Omron Sysmac Studio project AutomatedSortingSystem (Sysmac Studio 1.64.0.64008, StandardProject)

# Controller new_Controller_0: NJ301-1100 version 1.69
Units and slaves: Power Supply : NJ-Px3001; CPU : NJ301-1100
Task PrimaryTask (priority 4, period or condition 1000): PRG_SortingSystem

TYPE ST_MotorSimulation : STRUCT
    Enable : BOOL;
    Start : BOOL;
    Stop : BOOL;
    Fault : BOOL;
    RunFeedback : BOOL;
    ResetFault : BOOL;
    MotorRun : BOOL;
    MotorFault : BOOL;
    StartupFault : BOOL;
    FeedbackLostFault : BOOL;
END_STRUCT END_TYPE
TYPE ST_CylinderSimulation : STRUCT
    Enable : BOOL;
    ExtendCmd : BOOL;
    RetractCmd : BOOL;
    SensorExtended : BOOL;
    SensorRetracted : BOOL;
    ResetFault : BOOL;
    ValveExtend : BOOL;
    ValveRetract : BOOL;
    CylinderFault : BOOL;
    ExtendTimeoutFault : BOOL;
    RetractTimeoutFault : BOOL;
END_STRUCT END_TYPE
TYPE ST_SortingSimulation : STRUCT
    AutoMode : BOOL;
    Start : BOOL;
    Stop : BOOL;
    Reset : BOOL;
    ProductDetected : BOOL;
    AtSortingPosition : BOOL;
    ProductType : UINT;  (* 1=A, 2=B, 3=C *)
    CycleActive : BOOL;
    CycleComplete : BOOL;
    SystemFault : BOOL;
    ProductAtExit : BOOL;
END_STRUCT END_TYPE

PROGRAM Program0
VAR
    Motor1 : FB_ConveyorMotor;
    MotorSim : ST_MotorSimulation;
    CylinderSim : ST_CylinderSimulation;
    Cylinder1 : FB_PneumaticCylinder;
END_VAR

(* Section Section0: ladder, written here as Structured Text *)

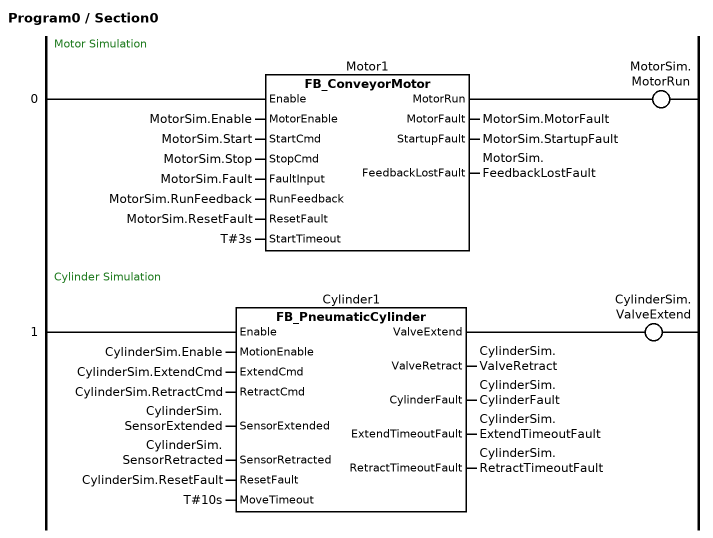
(* Rung 0: Motor Simulation *)
Motor1(Enable := TRUE, MotorEnable := MotorSim.Enable, StartCmd := MotorSim.Start, StopCmd := MotorSim.Stop, FaultInput := MotorSim.Fault, RunFeedback := MotorSim.RunFeedback, ResetFault := MotorSim.ResetFault, StartTimeout := T#3s, MotorFault => MotorSim.MotorFault, StartupFault => MotorSim.StartupFault, FeedbackLostFault => MotorSim.FeedbackLostFault);
MotorSim.MotorRun := Motor1.MotorRun;
(* Rung 1: Cylinder Simulation *)
Cylinder1(Enable := TRUE, MotionEnable := CylinderSim.Enable, ExtendCmd := CylinderSim.ExtendCmd, RetractCmd := CylinderSim.RetractCmd, SensorExtended := CylinderSim.SensorExtended, SensorRetracted := CylinderSim.SensorRetracted, ResetFault := CylinderSim.ResetFault, MoveTimeout := T#10s, ValveRetract => CylinderSim.ValveRetract, CylinderFault => CylinderSim.CylinderFault, ExtendTimeoutFault => CylinderSim.ExtendTimeoutFault, RetractTimeoutFault => CylinderSim.RetractTimeoutFault);
CylinderSim.ValveExtend := Cylinder1.ValveExtend;
END_PROGRAM

PROGRAM PRG_SortingSystem
VAR
    Motor_Conv1 : FB_ConveyorMotor;
    Motor_Conv2 : FB_ConveyorMotor;
    Motor_Conv3 : FB_ConveyorMotor;
    Cylinder_A : FB_PneumaticCylinder;
    Cylinder_B : FB_PneumaticCylinder;
    Conv1 : ST_MotorSimulation;
    Conv2 : ST_MotorSimulation;
    Conv3 : ST_MotorSimulation;
    CylA : ST_CylinderSimulation;
    CylB : ST_CylinderSimulation;
    SortingSim : ST_SortingSimulation;
    TestInput : BOOL;
    TestOutput : BOOL;
    SortingSequence : FB_SortingSequence;
    DevicesReady : BOOL;
    AnyDeviceFault : BOOL;
    SortingState : UINT;
    SystemEnable : BOOL;
    CylinderSim_A : FB_CylinderSimulator;
    CylinderSim_B : FB_CylinderSimulator;
    SimulateCylinderAJam : BOOL := False;
    SimulateCylinderBJam : BOOL := False;
    ResetCylinderAPosition : BOOL := False;
    ResetCylinderBPosition : BOOL := False;
    AlarmManager : FB_AlarmManager;
    ActiveAlarmCode : UINT;
    AlarmActiveStatus : BOOL;
END_VAR

(* Section Section0: ladder, written here as Structured Text *)

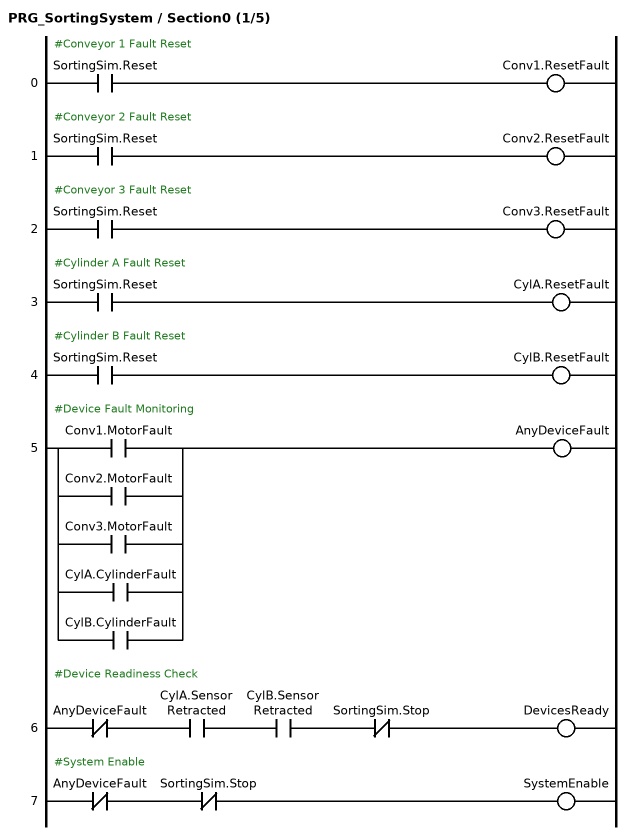
(* Rung 0: #Conveyor 1 Fault Reset *)
Conv1.ResetFault := SortingSim.Reset;
(* Rung 1: #Conveyor 2 Fault Reset *)
Conv2.ResetFault := SortingSim.Reset;
(* Rung 2: #Conveyor 3 Fault Reset *)
Conv3.ResetFault := SortingSim.Reset;
(* Rung 3: #Cylinder A Fault Reset *)
CylA.ResetFault := SortingSim.Reset;
(* Rung 4: #Cylinder B Fault Reset *)
CylB.ResetFault := SortingSim.Reset;
(* Rung 5: #Device Fault Monitoring *)
AnyDeviceFault := Conv1.MotorFault OR Conv2.MotorFault OR Conv3.MotorFault OR CylA.CylinderFault OR CylB.CylinderFault;
(* Rung 6: #Device Readiness Check *)
DevicesReady := NOT AnyDeviceFault AND CylA.SensorRetracted AND CylB.SensorRetracted AND NOT SortingSim.Stop;
(* Rung 7: #System Enable *)
SystemEnable := NOT AnyDeviceFault AND NOT SortingSim.Stop;

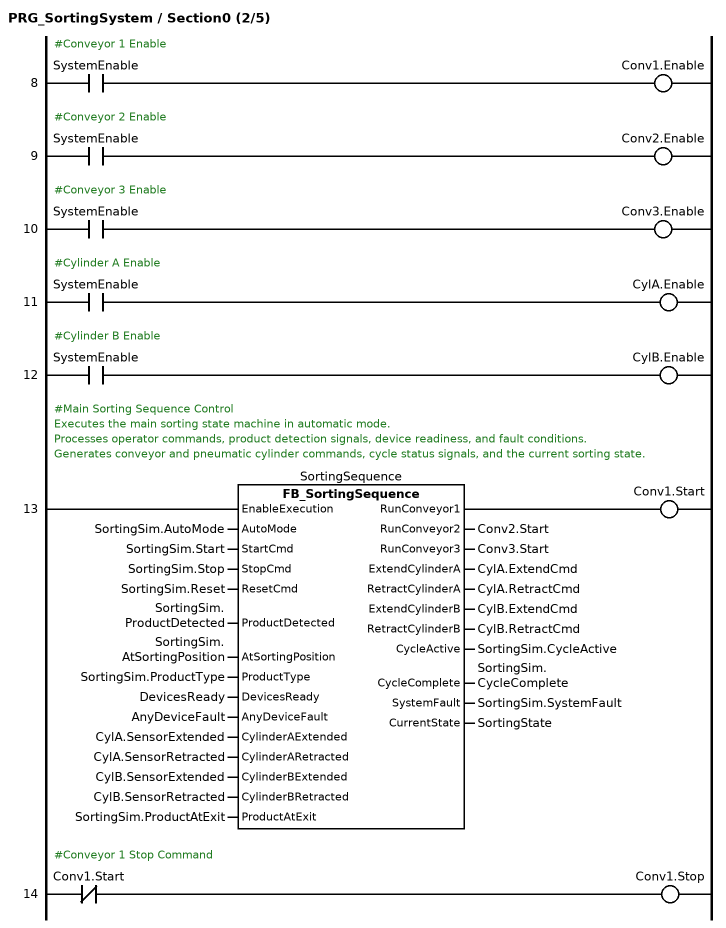
(* Rung 8: #Conveyor 1 Enable *)
Conv1.Enable := SystemEnable;
(* Rung 9: #Conveyor 2 Enable *)
Conv2.Enable := SystemEnable;
(* Rung 10: #Conveyor 3 Enable *)
Conv3.Enable := SystemEnable;
(* Rung 11: #Cylinder A Enable *)
CylA.Enable := SystemEnable;
(* Rung 12: #Cylinder B Enable *)
CylB.Enable := SystemEnable;
(* Rung 13: #Main Sorting Sequence Control / Executes the main sorting state machine in automatic mode. / Processes operator commands, product detection signals, device readiness, and fault conditions. / Generates conveyor and pneumatic cylinder commands, cycle status signals, and the current sorting state. *)
SortingSequence(EnableExecution := TRUE, AutoMode := SortingSim.AutoMode, StartCmd := SortingSim.Start, StopCmd := SortingSim.Stop, ResetCmd := SortingSim.Reset, ProductDetected := SortingSim.ProductDetected, AtSortingPosition := SortingSim.AtSortingPosition, ProductType := SortingSim.ProductType, DevicesReady := DevicesReady, AnyDeviceFault := AnyDeviceFault, CylinderAExtended := CylA.SensorExtended, CylinderARetracted := CylA.SensorRetracted, CylinderBExtended := CylB.SensorExtended, CylinderBRetracted := CylB.SensorRetracted, ProductAtExit := SortingSim.ProductAtExit, RunConveyor2 => Conv2.Start, RunConveyor3 => Conv3.Start, ExtendCylinderA => CylA.ExtendCmd, RetractCylinderA => CylA.RetractCmd, ExtendCylinderB => CylB.ExtendCmd, RetractCylinderB => CylB.RetractCmd, CycleActive => SortingSim.CycleActive, CycleComplete => SortingSim.CycleComplete, SystemFault => SortingSim.SystemFault, CurrentState => SortingState);
Conv1.Start := SortingSequence.RunConveyor1;
(* Rung 14: #Conveyor 1 Stop Command *)
Conv1.Stop := NOT Conv1.Start;

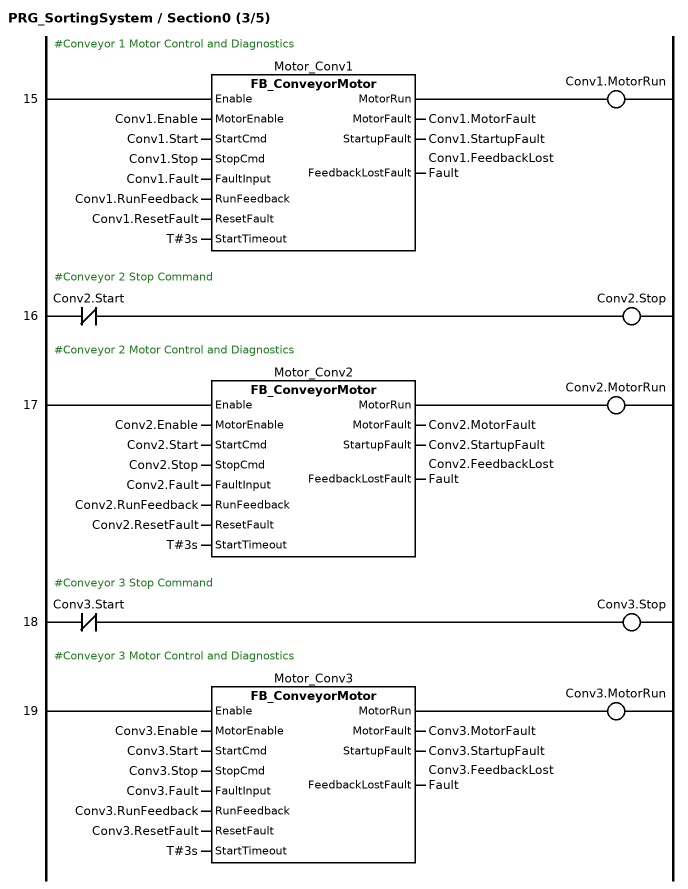
(* Rung 15: #Conveyor 1 Motor Control and Diagnostics *)
Motor_Conv1(Enable := TRUE, MotorEnable := Conv1.Enable, StartCmd := Conv1.Start, StopCmd := Conv1.Stop, FaultInput := Conv1.Fault, RunFeedback := Conv1.RunFeedback, ResetFault := Conv1.ResetFault, StartTimeout := T#3s, MotorFault => Conv1.MotorFault, StartupFault => Conv1.StartupFault, FeedbackLostFault => Conv1.FeedbackLostFault);
Conv1.MotorRun := Motor_Conv1.MotorRun;
(* Rung 16: #Conveyor 2 Stop Command *)
Conv2.Stop := NOT Conv2.Start;
(* Rung 17: #Conveyor 2 Motor Control and Diagnostics *)
Motor_Conv2(Enable := TRUE, MotorEnable := Conv2.Enable, StartCmd := Conv2.Start, StopCmd := Conv2.Stop, FaultInput := Conv2.Fault, RunFeedback := Conv2.RunFeedback, ResetFault := Conv2.ResetFault, StartTimeout := T#3s, MotorFault => Conv2.MotorFault, StartupFault => Conv2.StartupFault, FeedbackLostFault => Conv2.FeedbackLostFault);
Conv2.MotorRun := Motor_Conv2.MotorRun;
(* Rung 18: #Conveyor 3 Stop Command *)
Conv3.Stop := NOT Conv3.Start;
(* Rung 19: #Conveyor 3 Motor Control and Diagnostics *)
Motor_Conv3(Enable := TRUE, MotorEnable := Conv3.Enable, StartCmd := Conv3.Start, StopCmd := Conv3.Stop, FaultInput := Conv3.Fault, RunFeedback := Conv3.RunFeedback, ResetFault := Conv3.ResetFault, StartTimeout := T#3s, MotorFault => Conv3.MotorFault, StartupFault => Conv3.StartupFault, FeedbackLostFault => Conv3.FeedbackLostFault);
Conv3.MotorRun := Motor_Conv3.MotorRun;

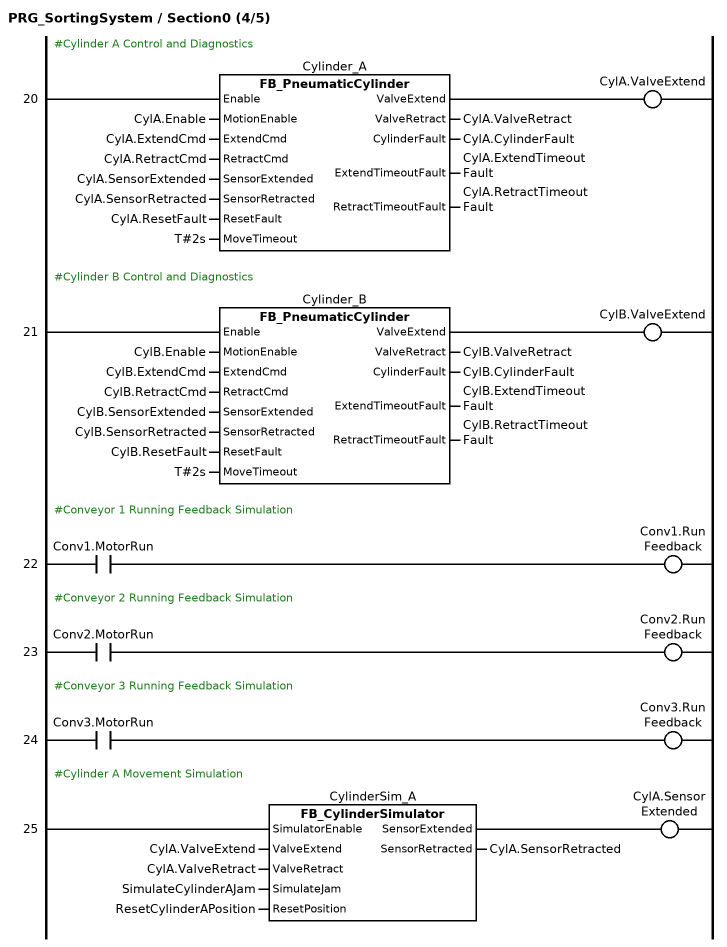
(* Rung 20: #Cylinder A Control and Diagnostics *)
Cylinder_A(Enable := TRUE, MotionEnable := CylA.Enable, ExtendCmd := CylA.ExtendCmd, RetractCmd := CylA.RetractCmd, SensorExtended := CylA.SensorExtended, SensorRetracted := CylA.SensorRetracted, ResetFault := CylA.ResetFault, MoveTimeout := T#2s, ValveRetract => CylA.ValveRetract, CylinderFault => CylA.CylinderFault, ExtendTimeoutFault => CylA.ExtendTimeoutFault, RetractTimeoutFault => CylA.RetractTimeoutFault);
CylA.ValveExtend := Cylinder_A.ValveExtend;
(* Rung 21: #Cylinder B Control and Diagnostics *)
Cylinder_B(Enable := TRUE, MotionEnable := CylB.Enable, ExtendCmd := CylB.ExtendCmd, RetractCmd := CylB.RetractCmd, SensorExtended := CylB.SensorExtended, SensorRetracted := CylB.SensorRetracted, ResetFault := CylB.ResetFault, MoveTimeout := T#2s, ValveRetract => CylB.ValveRetract, CylinderFault => CylB.CylinderFault, ExtendTimeoutFault => CylB.ExtendTimeoutFault, RetractTimeoutFault => CylB.RetractTimeoutFault);
CylB.ValveExtend := Cylinder_B.ValveExtend;
(* Rung 22: #Conveyor 1 Running Feedback Simulation *)
Conv1.RunFeedback := Conv1.MotorRun;
(* Rung 23: #Conveyor 2 Running Feedback Simulation *)
Conv2.RunFeedback := Conv2.MotorRun;
(* Rung 24: #Conveyor 3 Running Feedback Simulation *)
Conv3.RunFeedback := Conv3.MotorRun;
(* Rung 25: #Cylinder A Movement Simulation *)
CylinderSim_A(SimulatorEnable := TRUE, ValveExtend := CylA.ValveExtend, ValveRetract := CylA.ValveRetract, SimulateJam := SimulateCylinderAJam, ResetPosition := ResetCylinderAPosition, SensorRetracted => CylA.SensorRetracted);
CylA.SensorExtended := CylinderSim_A.SensorExtended;

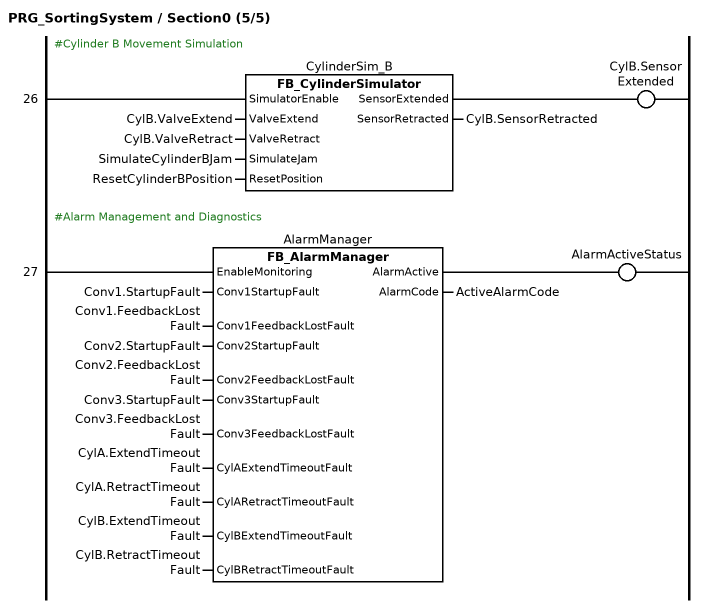
(* Rung 26: #Cylinder B Movement Simulation *)
CylinderSim_B(SimulatorEnable := TRUE, ValveExtend := CylB.ValveExtend, ValveRetract := CylB.ValveRetract, SimulateJam := SimulateCylinderBJam, ResetPosition := ResetCylinderBPosition, SensorRetracted => CylB.SensorRetracted);
CylB.SensorExtended := CylinderSim_B.SensorExtended;
(* Rung 27: #Alarm Management and Diagnostics *)
AlarmManager(EnableMonitoring := TRUE, Conv1StartupFault := Conv1.StartupFault, Conv1FeedbackLostFault := Conv1.FeedbackLostFault, Conv2StartupFault := Conv2.StartupFault, Conv2FeedbackLostFault := Conv2.FeedbackLostFault, Conv3StartupFault := Conv3.StartupFault, Conv3FeedbackLostFault := Conv3.FeedbackLostFault, CylAExtendTimeoutFault := CylA.ExtendTimeoutFault, CylARetractTimeoutFault := CylA.RetractTimeoutFault, CylBExtendTimeoutFault := CylB.ExtendTimeoutFault, CylBRetractTimeoutFault := CylB.RetractTimeoutFault, AlarmCode => ActiveAlarmCode);
AlarmActiveStatus := AlarmManager.AlarmActive;
END_PROGRAM

FUNCTION_BLOCK FB_ConveyorMotor
VAR
    StartTimer : TON;
    FaultLatch : BOOL;
    StartRequest : BOOL;
    StartCmdPrev : BOOL;
    StartEdge : BOOL;
    FeedbackTimer : TON;
    RunConfirmed : BOOL;
    StartupFaultLatch : BOOL;
    FeedbackFaultLatch : BOOL;
END_VAR
VAR_INPUT
    Enable : BOOL;
    MotorEnable : BOOL;
    StartCmd : BOOL;
    StopCmd : BOOL;
    FaultInput : BOOL;
    RunFeedback : BOOL;
    ResetFault : BOOL;
    StartTimeout : TIME := T#3s;
END_VAR
VAR_OUTPUT
    MotorRun : BOOL;
    MotorFault : BOOL;
    StartupFault : BOOL;
    FeedbackLostFault : BOOL;
END_VAR
//Detect rising edge of Start command
StartEdge := StartCmd AND NOT StartCmdPrev;
StartCmdPrev := StartCmd;

//Reset fault memory
IF ResetFault
   AND StopCmd
   AND NOT StartCmd
   AND NOT FaultInput THEN

    FaultLatch := FALSE;
    StartupFaultLatch := FALSE;
    FeedbackFaultLatch := FALSE;

END_IF;

//Accept a new Start command
IF StartEdge AND MotorEnable AND NOT StopCmd
   AND NOT FaultInput AND NOT FaultLatch THEN
    StartRequest := TRUE;
    RunConfirmed := FALSE;
END_IF;

//Stop and interlock handling
IF StopCmd OR NOT MotorEnable OR FaultInput OR FaultLatch THEN
    StartRequest := FALSE;
END_IF;

//Reset confirmation after stop
IF NOT StartRequest THEN
    RunConfirmed := FALSE;
END_IF;

//Motor command
MotorRun := StartRequest AND MotorEnable
            AND NOT StopCmd
            AND NOT FaultInput
            AND NOT FaultLatch;

//Remember successful start
IF MotorRun AND RunFeedback THEN
    RunConfirmed := TRUE;
END_IF;

//Startup timeout
StartTimer(
    IN := MotorRun AND NOT RunConfirmed,
    PT := StartTimeout
);

IF StartTimer.Q THEN
    StartupFaultLatch := TRUE;
    FaultLatch := TRUE;
END_IF;

//Feedback loss during operation
FeedbackTimer(
    IN := MotorRun AND RunConfirmed
          AND NOT RunFeedback,
    PT := T#1s
);

IF FeedbackTimer.Q THEN
    FeedbackFaultLatch := TRUE;
    FaultLatch := TRUE;
END_IF;

//Remove motor command on fault
IF FaultLatch THEN
    StartRequest := FALSE;
    MotorRun := FALSE;
    RunConfirmed := FALSE;
END_IF;

//Diagnostic outputs
StartupFault := StartupFaultLatch;
FeedbackLostFault := FeedbackFaultLatch;
MotorFault := FaultInput OR FaultLatch;
END_FUNCTION_BLOCK

FUNCTION_BLOCK FB_PneumaticCylinder
VAR
    ExtendTimer : TON;
    RetractTimer : TON;
    ExtendFaultLatch : BOOL;
    RetractFaultLatch : BOOL;
    SensorConflictLatch : BOOL;
END_VAR
VAR_INPUT
    Enable : BOOL;
    MotionEnable : BOOL;
    ExtendCmd : BOOL;
    RetractCmd : BOOL;
    SensorExtended : BOOL;
    SensorRetracted : BOOL;
    ResetFault : BOOL;
    MoveTimeout : TIME;
END_VAR
VAR_OUTPUT
    ValveExtend : BOOL;
    ValveRetract : BOOL;
    CylinderFault : BOOL;
    ExtendTimeoutFault : BOOL;
    RetractTimeoutFault : BOOL;
END_VAR
//Reset stored faults only when idle
IF ResetFault
   AND NOT ExtendCmd
   AND NOT RetractCmd
   AND NOT (SensorExtended AND SensorRetracted) THEN

    ExtendFaultLatch := FALSE;
    RetractFaultLatch := FALSE;
    SensorConflictLatch := FALSE;

END_IF;

//Detect contradictory position sensors
IF SensorExtended AND SensorRetracted THEN
    SensorConflictLatch := TRUE;
END_IF;

//General fault condition
CylinderFault := ExtendFaultLatch
                 OR RetractFaultLatch
                 OR SensorConflictLatch;

//Control valve outputs
ValveExtend := MotionEnable
               AND ExtendCmd
               AND NOT RetractCmd
               AND NOT SensorExtended
               AND NOT CylinderFault;

ValveRetract := MotionEnable
                AND RetractCmd
                AND NOT ExtendCmd
                AND NOT SensorRetracted
                AND NOT CylinderFault;

//Monitor extension movement
ExtendTimer(
    IN := ValveExtend AND NOT SensorExtended,
    PT := MoveTimeout
);

IF ExtendTimer.Q THEN
    ExtendFaultLatch := TRUE;
END_IF;

//Monitor retraction movement
RetractTimer(
    IN := ValveRetract AND NOT SensorRetracted,
    PT := MoveTimeout
);

IF RetractTimer.Q THEN
    RetractFaultLatch := TRUE;
END_IF;

//Update diagnostic outputs
ExtendTimeoutFault := ExtendFaultLatch;
RetractTimeoutFault := RetractFaultLatch;

CylinderFault := ExtendFaultLatch
                 OR RetractFaultLatch
                 OR SensorConflictLatch;

//Remove valve commands on fault
IF CylinderFault THEN
    ValveExtend := FALSE;
    ValveRetract := FALSE;
END_IF;
END_FUNCTION_BLOCK

FUNCTION_BLOCK FB_SortingSequence
VAR
    State : UINT;
    SelectedProduct : UINT;
    StartPrev : BOOL;
    StartEdge : BOOL;
    FaultLatch : BOOL;
    ExitSensorTriggered : BOOL;
    SortingPositionCleared : BOOL;
    ProductSensorReady : BOOL;
END_VAR
VAR_INPUT
    EnableExecution : BOOL;
    AutoMode : BOOL;
    StartCmd : BOOL;
    StopCmd : BOOL;
    ResetCmd : BOOL;
    ProductDetected : BOOL;
    AtSortingPosition : BOOL;
    ProductType : UINT;
    DevicesReady : BOOL;
    AnyDeviceFault : BOOL;
END_VAR
VAR_OUTPUT
    RunConveyor1 : BOOL;
    RunConveyor2 : BOOL;
    RunConveyor3 : BOOL;
    ExtendCylinderA : BOOL;
    RetractCylinderA : BOOL;
    ExtendCylinderB : BOOL;
    RetractCylinderB : BOOL;
    CycleActive : BOOL;
    CycleComplete : BOOL;
    SystemFault : BOOL;
    CurrentState : UINT;
END_VAR
VAR_INPUT
    CylinderAExtended : BOOL;
    CylinderARetracted : BOOL;
    CylinderBExtended : BOOL;
    CylinderBRetracted : BOOL;
    ProductAtExit : BOOL;
END_VAR
//Detect a new Start press
StartEdge := StartCmd AND NOT StartPrev;
StartPrev := StartCmd;

//Ignore Start while Stop, Reset or Fault is active
IF NOT EnableExecution OR StopCmd OR ResetCmd 
	OR NOT AutoMode OR FaultLatch OR AnyDeviceFault THEN
    StartEdge := FALSE;
END_IF;

//Default outputs
RunConveyor1 := FALSE;
RunConveyor2 := FALSE;
RunConveyor3 := FALSE;

ExtendCylinderA := FALSE;
RetractCylinderA := FALSE;
ExtendCylinderB := FALSE;
RetractCylinderB := FALSE;

CycleActive := FALSE;
CycleComplete := FALSE;

//Fault handling
IF AnyDeviceFault THEN
    FaultLatch := TRUE;
END_IF;

IF FaultLatch THEN
    State := UINT#900;
END_IF;

//Stop / Manual mode / Execution disabled
IF StopCmd OR NOT AutoMode OR NOT EnableExecution THEN
	ExitSensorTriggered := FALSE;
	SortingPositionCleared := FALSE;
	ProductSensorReady := FALSE;
	
    IF NOT FaultLatch THEN
        State := UINT#0;
        SelectedProduct := UINT#0;
    END_IF;
END_IF;

//Reset fault
IF ResetCmd
   AND NOT StartCmd
   AND NOT AnyDeviceFault THEN

    FaultLatch := FALSE;
    State := UINT#0;
    SelectedProduct := UINT#0;
	ExitSensorTriggered := FALSE;
	SortingPositionCleared := FALSE;
	ProductSensorReady := FALSE;

END_IF;

//Main state machine
IF EnableExecution
   AND AutoMode
   AND NOT StopCmd
   AND NOT ResetCmd
   AND NOT FaultLatch
   AND NOT AnyDeviceFault THEN
   
	CASE State OF

	    UINT#0: //IDLE
		    ExitSensorTriggered := FALSE;
		    SortingPositionCleared := FALSE;
		    ProductSensorReady := FALSE;

		    IF StartEdge AND DevicesReady THEN
		        SelectedProduct := UINT#0;
		        State := UINT#10;
		    END_IF;

	    UINT#10: //WAIT_FOR_PRODUCT
		    CycleActive := TRUE;
		    RunConveyor1 := TRUE;
		    RunConveyor2 := TRUE;
		    RunConveyor3 := TRUE;

	    	//Confirm that sorting position is clear
		    IF NOT AtSortingPosition THEN
		        SortingPositionCleared := TRUE;
		    END_IF;
			
			//Arm product detection after sensor is released
		    IF NOT ProductDetected THEN
		        ProductSensorReady := TRUE;
		    END_IF;

	    	//Accept a new product only when position is clear
		    IF ProductDetected AND ProductSensorReady AND SortingPositionCleared THEN
		        SelectedProduct := ProductType;
				ProductSensorReady := FALSE;
		        State := UINT#20;
		    END_IF;

	    UINT#20: //TRANSPORT
	        CycleActive := TRUE;
	        RunConveyor1 := TRUE;
	        RunConveyor2 := TRUE;
	        RunConveyor3 := TRUE;

	        IF AtSortingPosition AND SortingPositionCleared THEN
	    		SortingPositionCleared := FALSE;
				
	            CASE SelectedProduct OF
	                UINT#1:
	                    State := UINT#30;
	                UINT#2:
	                    State := UINT#40;
	                UINT#3:
	                    State := UINT#50;
	                ELSE
	                    FaultLatch := TRUE;
	                    State := UINT#900;
	            END_CASE;
	        END_IF;

	    UINT#30: //EXTEND_A
	        CycleActive := TRUE;
	        RunConveyor2 := TRUE;
	        ExtendCylinderA := TRUE;

	        IF CylinderAExtended THEN
	            State := UINT#31;
	        END_IF;

	    UINT#31: //RETRACT_A
	        CycleActive := TRUE;
	        RunConveyor2 := TRUE;
	        RetractCylinderA := TRUE;

	        IF CylinderARetracted THEN
	            State := UINT#60;
	        END_IF;

	    UINT#40: //EXTEND_B
	        CycleActive := TRUE;
	        RunConveyor3 := TRUE;
	        ExtendCylinderB := TRUE;

	        IF CylinderBExtended THEN
	            State := UINT#41;
	        END_IF;

	    UINT#41: //RETRACT_B
	        CycleActive := TRUE;
	        RunConveyor3 := TRUE;
	        RetractCylinderB := TRUE;

	        IF CylinderBRetracted THEN
	            State := UINT#60;
	        END_IF;
	    
		UINT#50: //SORT_C
		    CycleActive := TRUE;
		    RunConveyor1 := TRUE;

		    //Wait until exit sensor is clear
		    IF NOT ProductAtExit THEN
		        ExitSensorTriggered := FALSE;
		        State := UINT#51;
		    END_IF;

		UINT#51: //WAIT_EXIT_DETECTION
		    CycleActive := TRUE;
		    RunConveyor1 := TRUE;

		    IF ProductAtExit THEN
		        ExitSensorTriggered := TRUE;
		        State := UINT#52;
		    END_IF;

		UINT#52: //WAIT_EXIT_CLEAR
		    CycleActive := TRUE;
		    RunConveyor1 := TRUE;

		    IF ExitSensorTriggered AND NOT ProductAtExit THEN
		        ExitSensorTriggered := FALSE;
		        State := UINT#60;
		    END_IF;


	    UINT#60: //COMPLETE
	        CycleComplete := TRUE;
	        State := UINT#10;

	    UINT#900: //FAULT
	        ; //Fault state - outputs are handled by the final interlock

	    ELSE
	        State := UINT#0;

	END_CASE;
	
END_IF;

//Final output interlock
IF NOT EnableExecution
   OR StopCmd OR ResetCmd OR NOT AutoMode
   OR FaultLatch OR AnyDeviceFault THEN
    RunConveyor1 := FALSE;
    RunConveyor2 := FALSE;
    RunConveyor3 := FALSE;

    ExtendCylinderA := FALSE;
    RetractCylinderA := FALSE;
    ExtendCylinderB := FALSE;
    RetractCylinderB := FALSE;

    CycleActive := FALSE;
    CycleComplete := FALSE;
END_IF;

//Diagnostic outputs
CurrentState := State;
SystemFault := FaultLatch;
END_FUNCTION_BLOCK

FUNCTION_BLOCK FB_CylinderSimulator
VAR
    ExtendDelay : TON;
    RetractDelay : TON;
    Position : UINT := 0;
END_VAR
VAR_INPUT
    SimulatorEnable : BOOL;
    ValveExtend : BOOL;
    ValveRetract : BOOL;
END_VAR
VAR_OUTPUT
    SensorExtended : BOOL;
    SensorRetracted : BOOL;
END_VAR
VAR_INPUT
    SimulateJam : BOOL := False;
    ResetPosition : BOOL := False;
END_VAR
//Cylinder movement simulation
ExtendDelay(
    IN := ValveExtend AND NOT ValveRetract AND NOT SimulateJam,
    PT := T#500ms
);

RetractDelay(
    IN := ValveRetract AND NOT ValveExtend AND NOT SimulateJam,
    PT := T#500ms
);

IF ExtendDelay.Q THEN
    Position := UINT#2;
ELSIF RetractDelay.Q THEN
    Position := UINT#0;
ELSIF ValveExtend AND NOT ValveRetract THEN
    Position := UINT#1;
ELSIF ValveRetract AND NOT ValveExtend THEN
    Position := UINT#1;
END_IF;

//Manual reset of simulated cylinder position
IF ResetPosition THEN
    Position := UINT#0;
END_IF;

//Simulated position sensors
SensorExtended := (Position = UINT#2);
SensorRetracted := (Position = UINT#0);
END_FUNCTION_BLOCK

FUNCTION_BLOCK FB_AlarmManager
VAR_INPUT
    EnableMonitoring : BOOL;
    Conv1StartupFault : BOOL;
    Conv1FeedbackLostFault : BOOL;
    Conv2StartupFault : BOOL;
    Conv2FeedbackLostFault : BOOL;
    Conv3StartupFault : BOOL;
    Conv3FeedbackLostFault : BOOL;
    CylAExtendTimeoutFault : BOOL;
    CylARetractTimeoutFault : BOOL;
    CylBExtendTimeoutFault : BOOL;
    CylBRetractTimeoutFault : BOOL;
END_VAR
VAR_OUTPUT
    AlarmActive : BOOL;
    AlarmCode : UINT;
END_VAR
//Default outputs
AlarmActive := FALSE;
AlarmCode := UINT#0;

IF EnableMonitoring THEN

    //Alarm selection based on priority
    IF Conv1StartupFault THEN
        AlarmCode := UINT#101;

    ELSIF Conv1FeedbackLostFault THEN
        AlarmCode := UINT#102;

    ELSIF Conv2StartupFault THEN
        AlarmCode := UINT#201;

    ELSIF Conv2FeedbackLostFault THEN
        AlarmCode := UINT#202;

    ELSIF Conv3StartupFault THEN
        AlarmCode := UINT#301;

    ELSIF Conv3FeedbackLostFault THEN
        AlarmCode := UINT#302;

    ELSIF CylAExtendTimeoutFault THEN
        AlarmCode := UINT#401;

    ELSIF CylARetractTimeoutFault THEN
        AlarmCode := UINT#402;

    ELSIF CylBExtendTimeoutFault THEN
        AlarmCode := UINT#501;

    ELSIF CylBRetractTimeoutFault THEN
        AlarmCode := UINT#502;
    END_IF;

    //Alarm status
    AlarmActive := (AlarmCode <> UINT#0);

END_IF;
END_FUNCTION_BLOCK